Fanuc KAREL source: kb00154.KL

PROGRAM KB00154
%STACKSIZE=65535
%PRIORITY=65535
%NOLOCKGROUP
VAR
P1 : STRING[80]
P2 : STRING[80]
P3 : INTEGER
BEGIN
P1='A'
P2='A'
P3=1
SAVE(P1,P2,P3,1)
END KB00154
